(* IEC 61131-3 sources: plc-vscode/tests/st/test-ready/trust-platform/examples/OSCAT/cooling_tower_facade_template/non-oop/src, 3 files *)

(* ---- Main.st ---- *)
FUNCTION_BLOCK ClassicCoolingTower
VAR
    BasinHeaterValue : BOOL;
    BleedValveValue : BOOL;
    SeasonIdValue : INT;
END_VAR
METHOD PUBLIC Update : INT
VAR_INPUT
    SeasonRequest : INT;
    WaterTempC : REAL;
    OutdoorTempC : REAL;
    ConductivityUs : REAL;
END_VAR
VAR
    FanThreshold : REAL;
    FreezeThreshold : REAL;
END_VAR
IF SeasonRequest = INT#2 THEN
    SeasonIdValue := INT#2;
    FanThreshold := REAL#32.0;
    FreezeThreshold := REAL#4.0;
ELSE
    SeasonIdValue := INT#1;
    FanThreshold := REAL#26.0;
    FreezeThreshold := REAL#-10.0;
END_IF;
BasinHeaterValue := OutdoorTempC < FreezeThreshold;
BleedValveValue := ConductivityUs > REAL#1800.0;
IF WaterTempC > (FanThreshold + REAL#5.0) THEN
    Update := INT#2;
ELSIF WaterTempC > FanThreshold THEN
    Update := INT#1;
ELSE
    Update := INT#0;
END_IF;
END_METHOD
PUBLIC PROPERTY BasinHeater : BOOL
GET
    BasinHeater := BasinHeaterValue;
END_GET
END_PROPERTY
END_FUNCTION_BLOCK
PROGRAM Main
VAR
    Tower : ClassicCoolingTower;
    FanStage : INT;
END_VAR
FanStage := Tower.Update(SeasonRequest := INT#1, WaterTempC := REAL#32.0, OutdoorTempC := REAL#20.0, ConductivityUs := REAL#1000.0);
END_PROGRAM

(* ---- Configuration.st ---- *)
CONFIGURATION CoolingTowerFacadeTemplateClassicConfiguration
RESOURCE Cpu0 ON PLC
    TASK MainTask (INTERVAL := T#100ms, PRIORITY := 1);
    PROGRAM Tower WITH MainTask : Main;
END_RESOURCE
END_CONFIGURATION

(* ---- Tests.st ---- *)
TEST_PROGRAM ClassicCoolingTowerBranchesOnSeason
VAR
    Tower : ClassicCoolingTower;
END_VAR
ASSERT_EQUAL(EXPECTED := INT#2, ACTUAL := Tower.Update(SeasonRequest := INT#1, WaterTempC := REAL#32.0, OutdoorTempC := REAL#20.0, ConductivityUs := REAL#1000.0));
Tower.Update(SeasonRequest := INT#2, WaterTempC := REAL#20.0, OutdoorTempC := REAL#0.0, ConductivityUs := REAL#2000.0);
ASSERT_TRUE(IN := Tower.BasinHeater);
END_TEST_PROGRAM
